// TIA Portal project "Lamppu_saato" (V16)

(* hardware
DEVICE "Lamppuprosessi PLC 1200"  S7-1200 Station
   slot 0: "S7-1200 rack"  S7-1200 Rack  Rack  V1.0
   slot 1: "PLC5"  CPU 1214C DC/DC/DC  6ES7 214-1AG40-0XB0  V4.1
   slot 2: "AI 4xRTD_1"  SM 1231 AI4 x RTD  6ES7 231-5PD32-0XB0  V2.0
   slot 3: "AQ 1x12BIT_1"  AQ1 signal board  6ES7 232-4HA30-0XB0  V1.0
*)

// ===== PLC "PLC5"  CPU 1214C DC/DC/DC =====

VAR_GLOBAL   // PLC tag table "Default tag table"
   "bStart" AT %I0.0 : Bool;
   "iwPt100" AT %IW96 : Word;
   "Tag_1" AT %I2.0 : Bool;   // Ensimmäisen tulokortin 1 tulo
   "Tag_2" AT %I2.1 : Bool;
   "qwLamppu" AT %QW80 : Word;
   "bLaitepaalla" AT %Q0.0 : Bool;
   "Tag_3" AT %Q2.0 : Bool;   // Ensimmäisen lähtökortin 1 lähtö
   "Tag_4" AT %Q2.1 : Bool;
   "rLampoOlo" AT %MD100 : Real;
   "rLampoOhje" AT %MD104 : Real;
   "rPIDOutput" AT %MD108 : Real;
END_VAR

ORGANIZATION_BLOCK "Main"   // OB1, FBD, ProgramCycle
TITLE = "Main Program Sweep (Cycle)"
{ S7_Optimized_Access := 'TRUE' }
VERSION : 0.1
BEGIN

REGION Network 1
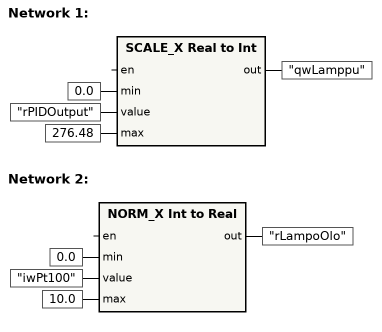
   "qwLamppu" := SCALE_X(MIN := 0.0, VALUE := "rPIDOutput", MAX := 276.48);
END_REGION

REGION Network 2
   "rLampoOlo" := NORM_X(MIN := 0.0, VALUE := "iwPt100", MAX := 10.0);
END_REGION
END_ORGANIZATION_BLOCK

ORGANIZATION_BLOCK "Cyclic interrupt"   // OB30, FBD, CyclicInterrupt
{ S7_Optimized_Access := 'TRUE' }
VERSION : 0.1
   VAR_INPUT
      Initial_Call : Bool;   // Initial call of this OB
      Event_Count : Int;   // Events discarded
   END_VAR
BEGIN

REGION Network 1
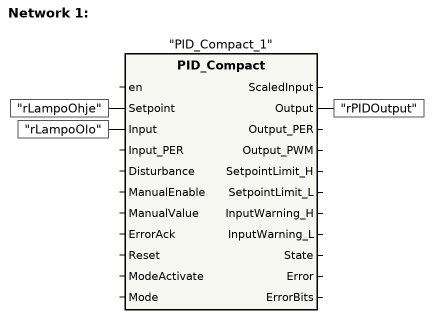
   "PID_Compact_1"(Setpoint := "rLampoOhje", Input := "rLampoOlo", Output => "rPIDOutput");   // PID_Compact
END_REGION
END_ORGANIZATION_BLOCK